(* IEC 61131-3 sources: trust-platform/examples/control/05-experiments-identification-and-validation/22-excitation-for-dynamics/src, 2 files *)

(* ---- Main.st ---- *)
(* Command of a periodic excitation about an operating point: u = u0 + d·sin(ω·t), with d in percentage points, ω in
   rad/s and t in s. *)
FUNCTION SineCommand : LREAL
VAR_INPUT
    OperatingPct : LREAL;
    AmplitudePct : LREAL;
    OmegaRadS : LREAL;
    ElapsedS : LREAL;
END_VAR
SineCommand := OperatingPct + AmplitudePct * SIN(OmegaRadS * ElapsedS);
END_FUNCTION

(* One heater's excitation: from Start, five periods P = 2π/ω of the sine about 75 %, then 75 % again. A setting
   outside 5–10 points or 0.05–1 rad/s is rejected and excites nothing; the command never leaves 0–100 %. *)
FUNCTION_BLOCK PeriodicExcitation
VAR_INPUT
    Start : BOOL;
    Enable : BOOL;
    AmplitudePct : LREAL;
    OmegaRadS : LREAL;
END_VAR
VAR_OUTPUT
    CommandPct : LREAL := 75.0;
    ElapsedS : LREAL := 0.0;
    Running : BOOL := FALSE;
    Rejected : BOOL := FALSE;
END_VAR
VAR
    OperatingPct : LREAL := 75.0;
    Periods : LREAL := 5.0;
    UpdateS : LREAL := 0.1;
END_VAR
Rejected := AmplitudePct < LREAL#5.0 OR AmplitudePct > LREAL#10.0 OR OmegaRadS < LREAL#0.05 OR OmegaRadS > LREAL#1.0;
IF Start AND NOT Rejected THEN
    Running := TRUE;
    ElapsedS := LREAL#0.0;
END_IF;
IF NOT Enable OR Rejected THEN
    Running := FALSE;
END_IF;
IF Running AND ElapsedS >= Periods * LREAL#2.0 * LREAL#3.14159265358979 / OmegaRadS - LREAL#1.0E-9 THEN
    Running := FALSE;
END_IF;
IF Running THEN
    CommandPct := LIMIT(LREAL#0.0, SineCommand(OperatingPct := OperatingPct, AmplitudePct := AmplitudePct,
        OmegaRadS := OmegaRadS, ElapsedS := ElapsedS), LREAL#100.0);
    ElapsedS := ElapsedS + UpdateS;
ELSE
    CommandPct := OperatingPct;
END_IF;
END_FUNCTION_BLOCK

PROGRAM Main
VAR
    (* Three copies of the heater at 35 °C, excited with the same amplitude at three rates. The heater control is
       off: the program sets the heater command directly. *)
    MiddleExcitation : PeriodicExcitation;
    SlowExcitation : PeriodicExcitation;
    FastExcitation : PeriodicExcitation;
    AmplitudePct : LREAL := 5.0;
    MiddleOmegaRadS : LREAL := 0.2;
    SlowOmegaRadS : LREAL := 0.1;
    FastOmegaRadS : LREAL := 0.4;
    MiddleTemperatureC : LREAL := 35.0;
    SlowTemperatureC : LREAL := 35.0;
    FastTemperatureC : LREAL := 35.0;
    MiddleCommandPct : LREAL := 75.0;
    SlowCommandPct : LREAL := 75.0;
    FastCommandPct : LREAL := 75.0;
    (* Control Studio's project experiment starts all three excitations at once. *)
    ExperimentEnabled : BOOL := FALSE;
    ExperimentWasEnabled : BOOL := FALSE;
    Start : BOOL := FALSE;
END_VAR

Start := ExperimentEnabled AND NOT ExperimentWasEnabled;
ExperimentWasEnabled := ExperimentEnabled;
MiddleExcitation(Start := Start, Enable := ExperimentEnabled, AmplitudePct := AmplitudePct, OmegaRadS := MiddleOmegaRadS);
SlowExcitation(Start := Start, Enable := ExperimentEnabled, AmplitudePct := AmplitudePct, OmegaRadS := SlowOmegaRadS);
FastExcitation(Start := Start, Enable := ExperimentEnabled, AmplitudePct := AmplitudePct, OmegaRadS := FastOmegaRadS);
MiddleCommandPct := MiddleExcitation.CommandPct;
SlowCommandPct := SlowExcitation.CommandPct;
FastCommandPct := FastExcitation.CommandPct;
END_PROGRAM

CONFIGURATION Config
RESOURCE Res ON PLC
    TASK MainTask(INTERVAL := T#100ms, PRIORITY := 1);
    PROGRAM P1 WITH MainTask : Main;
END_RESOURCE
VAR_CONFIG
    P1.MiddleCommandPct AT %QL0 : LREAL;
    P1.SlowCommandPct AT %QL8 : LREAL;
    P1.FastCommandPct AT %QL16 : LREAL;
    P1.MiddleTemperatureC AT %IL0 : LREAL;
    P1.SlowTemperatureC AT %IL8 : LREAL;
    P1.FastTemperatureC AT %IL16 : LREAL;
    P1.ExperimentEnabled AT %MX24.0 : BOOL;
END_VAR
END_CONFIGURATION

(* ---- tests.st ---- *)
(* @trustlsp:runtime-ignore — run these assertions with trust-dev test;
   they are not scheduled PLC instances in the lesson simulator. *)

TEST_PROGRAM TheSineAboutTheOperatingPoint
(* u = 75 + 5·sin(0.2·t): a period of 2π/0.2 = 31.416 s, 80 % a quarter period in, 70 % at three quarters. *)
ASSERT_NEAR(EXPECTED := LREAL#75.0, ACTUAL := SineCommand(OperatingPct := LREAL#75.0, AmplitudePct := LREAL#5.0,
    OmegaRadS := LREAL#0.2, ElapsedS := LREAL#0.0), DELTA := LREAL#1.0e-12);
ASSERT_NEAR(EXPECTED := LREAL#80.0, ACTUAL := SineCommand(OperatingPct := LREAL#75.0, AmplitudePct := LREAL#5.0,
    OmegaRadS := LREAL#0.2, ElapsedS := LREAL#7.853981633974483), DELTA := LREAL#1.0e-9);
ASSERT_NEAR(EXPECTED := LREAL#70.0, ACTUAL := SineCommand(OperatingPct := LREAL#75.0, AmplitudePct := LREAL#5.0,
    OmegaRadS := LREAL#0.2, ElapsedS := LREAL#23.56194490192345), DELTA := LREAL#1.0e-9);
END_TEST_PROGRAM

TEST_PROGRAM TheExcitationRunsFivePeriods
VAR
    Excitation : PeriodicExcitation;
    Updates : INT := 0;
    Count : INT;
END_VAR
(* ω = 0.4 rad/s: five periods are 78.54 s, 786 updates of 0.1 s; afterwards the command is 75 % again. *)
Excitation(Start := TRUE, Enable := TRUE, AmplitudePct := LREAL#5.0, OmegaRadS := LREAL#0.4);
IF Excitation.Running THEN
    Updates := 1;
END_IF;
FOR Count := 1 TO 900 DO
    Excitation(Start := FALSE, Enable := TRUE, AmplitudePct := LREAL#5.0, OmegaRadS := LREAL#0.4);
    IF Excitation.Running THEN
        Updates := Updates + 1;
    END_IF;
END_FOR;
ASSERT_EQUAL(EXPECTED := 786, ACTUAL := Updates);
ASSERT_NEAR(EXPECTED := LREAL#75.0, ACTUAL := Excitation.CommandPct, DELTA := LREAL#1.0e-12);
END_TEST_PROGRAM

TEST_PROGRAM ARejectedSettingExcitesNothing
VAR
    Excitation : PeriodicExcitation;
END_VAR
(* 20 points would drive the heater between 55 % and 95 %: outside the 5–10 points allowed here. *)
Excitation(Start := TRUE, Enable := TRUE, AmplitudePct := LREAL#20.0, OmegaRadS := LREAL#0.2);
ASSERT_TRUE(IN := Excitation.Rejected);
ASSERT_FALSE(IN := Excitation.Running);
ASSERT_NEAR(EXPECTED := LREAL#75.0, ACTUAL := Excitation.CommandPct, DELTA := LREAL#1.0e-12);
END_TEST_PROGRAM
